Fanuc KAREL source: kb00011.KL

PROGRAM KB00011
%NOLOCKGROUP
VAR
P1 : STRING[80];P2 : STRING[80];P3:INTEGER;P4:INTEGER;P5:INTEGER
BEGIN
--
--
--
--
P1='A'
P2='A'
P3=1
P4=1
P5=1
ATT_WINDOW_S(P1,P2,P3,P4,P5)
END KB00011
